// TIA Portal V21 export
// export: Created 2026-11-08T21:21:38.4892945Z, ExportSetting WithDefaults, DisplayName Totally Integrated Automation Portal, DisplayVersion V21 Update 3, DisplayName STEP 7 Professional, DisplayVersion V21 Update 3, DisplayName STEP 7 Safety, DisplayVersion V21, DisplayName Tech WebApplication, DisplayVersion V21, DisplayName WinCC Basic/Comfort/Advanced, DisplayVersion V21 Update 3, DisplayName WinCC Unified, DisplayVersion V21 Update 3
FUNCTION_BLOCK "FB_Stl"   // FB3, STL
TITLE = STL test FB
{ S7_Optimized_Access := 'TRUE' }
VERSION : 0.1
// stored: AutoNumber true, IsRetainMemResEnabled false, MemoryReserve 100, UDAEnableTagReadback false
   VAR_INPUT
      start : Bool;
      stop : Bool;
   END_VAR
   VAR_OUTPUT
      running : Bool;
      count : Int;
   END_VAR
   VAR
      cnt : Int;
      edge : Bool;
   END_VAR
BEGIN

NETWORK
TITLE = Latch
      A(;
      O     #start;
      O     #running;
      );
      AN    #stop;
      =     #running;

NETWORK
TITLE = Count rising edges
      A     #start;
      FP    #edge;
      JCN   END1;
      L     #cnt;
      +     1;
      T     #cnt;
END1: L     #cnt;
      T     #count;
      SET;
      SAVE;
END_FUNCTION_BLOCK
